TYPE ST_TcError :
STRUCT
	
	code 			: UDINT;
	message			: T_MaxString;
	
END_STRUCT
END_TYPE

(* stored: Version 1.1.0.1, ProductVersion 3.1.4024.12
   DUT ST_TcError: Id {b9a6efbd-1209-45d4-a4b5-cfdf5f94c984} *)
